PROGRAM POU_PBD
VAR
END_VAR

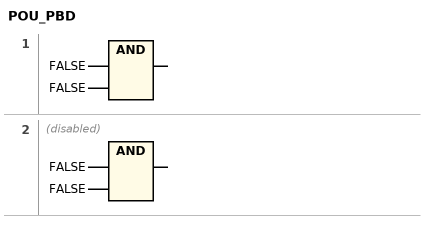
// NETWORK 1
(* FALSE AND FALSE; result not used *)

// NETWORK 2 (disabled)
// (* FALSE AND FALSE; result not used *)

END_PROGRAM

(* stored: Version 1.1.0.1, ProductVersion 3.1.4024.16
   POU POU_PBD: Id {60608d3c-cc8f-4eb3-9b00-632cb48a4b4b}, SpecialFunc None *)
